SUBAPPLICATION Uebung_094c_AX (* Zwei unabhaengige VT-Dropdowns (InputNumber_I1/I2) schalten je eine eigene Optionsgruppe frei: AD_TO_AUI -> AOption_AUI_DEMUX_1 -> OptionalGroup_001/002 per AOption-Adapter und QI. Noch OHNE gegenseitigen Ausschluss zwischen den beiden Gruppen - das braeuchte einen vorgeschalteten Arbiter, der aus den zwei unabhaengigen Dropdown-Events einen gemeinsamen K-Wert ableitet (offene Rueckfrage aus Krauternter: Bunker_Klappen/Aufnahme_Rechts, 'letzter Aktiviert gewinnt' + Boot-Tiebreak). *)
  (* Standard: 61499-2; Description: Copyright (c) 2026 Meisterschulen am Ostbahnhof This program and the accompanying materials are made available under the terms of the Eclipse Public License 2.0 which is available at https://www.eclipse.org/legal/epl-2.0/ SPDX-License-Identifier: EPL-2.0 *)
  (* Version 1.0, 2026-10-13, Franz Höpfinger, Meisterschulen am Ostbahnhof, initial API and implementation and/or initial documentation *)
  PACKAGE Uebungen;
  IMPORT Uebungen::const::UT::DefaultPool::InputNumber_I1;
  IMPORT Uebungen::const::UT::DefaultPool::InputNumber_I2;
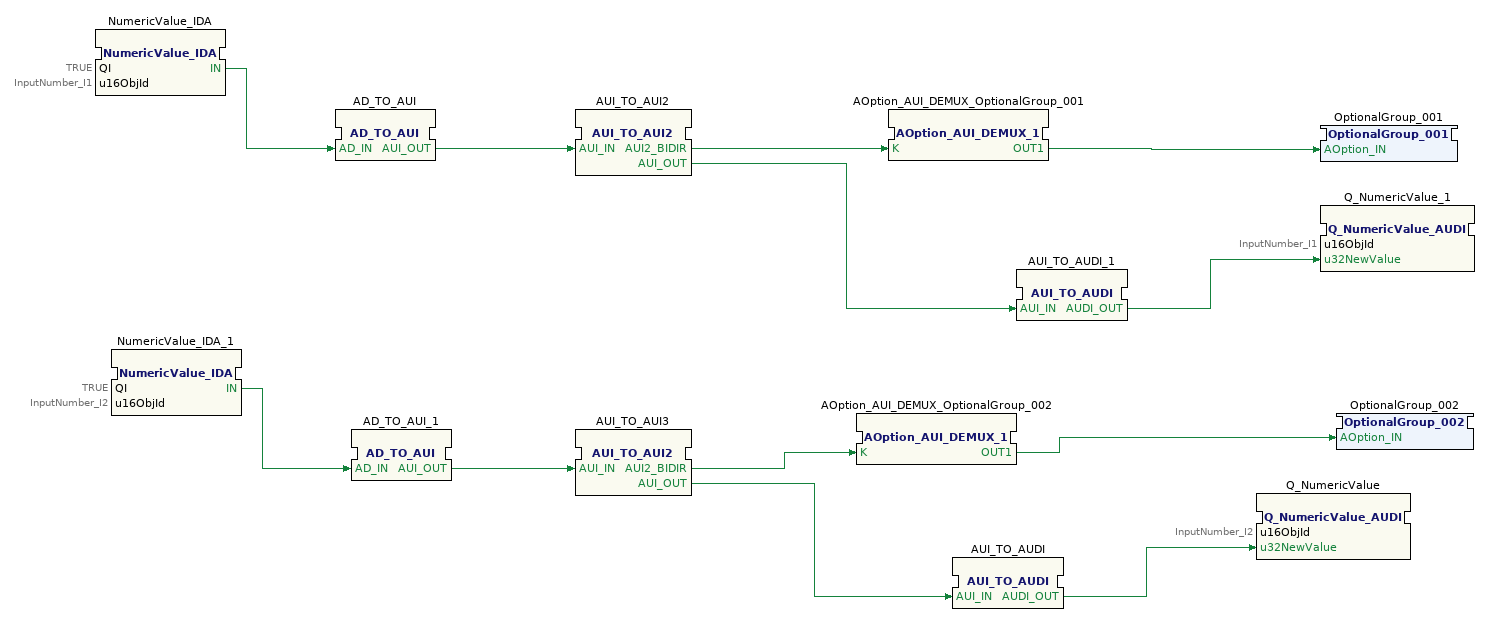
  FBS
    AOption_AUI_DEMUX_OptionalGroup_001 : Option::selection::AOption_AUI_DEMUX_1;
    NumericValue_IDA : isobus::UT::io::NumericValue::NumericValue_IDA(QI := TRUE, u16ObjId := InputNumber_I1);
    AD_TO_AUI : adapter::conversion::unidirectional::AD_TO_AUI;
    NumericValue_IDA_1 : isobus::UT::io::NumericValue::NumericValue_IDA(QI := TRUE, u16ObjId := InputNumber_I2);
    AOption_AUI_DEMUX_OptionalGroup_002 : Option::selection::AOption_AUI_DEMUX_1;
    AD_TO_AUI_1 : adapter::conversion::unidirectional::AD_TO_AUI;
    AUI_TO_AUI2 : adapter::conversion::bidirectional::AUI_TO_AUI2;
    AUI_TO_AUI3 : adapter::conversion::bidirectional::AUI_TO_AUI2;
    Q_NumericValue : isobus::UT::Q::Q_NumericValue_AUDI(u16ObjId := InputNumber_I2);
    AUI_TO_AUDI : adapter::conversion::unidirectional::AUI_TO_AUDI;
    AUI_TO_AUDI_1 : adapter::conversion::unidirectional::AUI_TO_AUDI;
    Q_NumericValue_1 : isobus::UT::Q::Q_NumericValue_AUDI(u16ObjId := InputNumber_I1);
  END_FBS
  SUBAPPS
    OptionalGroup_001 : MyLib_AX_Option::sys::OptionalGroup_001;
    OptionalGroup_002 : MyLib_AX_Option::sys::OptionalGroup_002;
  END_SUBAPPS
  ADAPTER_CONNECTIONS
    NumericValue_IDA.IN TO AD_TO_AUI.AD_IN;
    AD_TO_AUI.AUI_OUT TO AUI_TO_AUI2.AUI_IN;
    AOption_AUI_DEMUX_OptionalGroup_001.OUT1 TO OptionalGroup_001.AOption_IN;
    NumericValue_IDA_1.IN TO AD_TO_AUI_1.AD_IN;
    AOption_AUI_DEMUX_OptionalGroup_002.OUT1 TO OptionalGroup_002.AOption_IN;
    AUI_TO_AUI2.AUI2_BIDIR TO AOption_AUI_DEMUX_OptionalGroup_001.K;
    AD_TO_AUI_1.AUI_OUT TO AUI_TO_AUI3.AUI_IN;
    AUI_TO_AUI3.AUI2_BIDIR TO AOption_AUI_DEMUX_OptionalGroup_002.K;
    AUI_TO_AUDI.AUDI_OUT TO Q_NumericValue.u32NewValue;
    AUI_TO_AUI3.AUI_OUT TO AUI_TO_AUDI.AUI_IN;
    AUI_TO_AUDI_1.AUDI_OUT TO Q_NumericValue_1.u32NewValue;
    AUI_TO_AUI2.AUI_OUT TO AUI_TO_AUDI_1.AUI_IN;
  END_CONNECTIONS
END_SUBAPPLICATION
